FUNCTION_BLOCK Thomas_Object EXTENDS TcoCore.TcoObject
VAR
	_frank 		:	AKid_Object(THIS^);
	_andrew 	:	AKid_Object(THIS^);
	_christina 	:	AKid_Object(THIS^);
	_gianna 	:	AKid_Object(THIS^);
END_VAR

VAR
	_AskForTheFavor			:	AskForTheFavor_Task(THIS^);
END_VAR

METHOD AskForTheFavor : TcoCore.ITcoTask
VAR_INPUT
	Person_Requested 	:	REFERENCE TO Person_Object;
	RequestedFavor		:	STRING;
	ReturnFavor			:	STRING;
END_VAR
_AskForTheFavor(_Person_Requested := Person_Requested,_RequestedFavor :=RequestedFavor,_ReturnFavor:=ReturnFavor);

AskForTheFavor := _AskForTheFavor;
END_METHOD

END_FUNCTION_BLOCK

(* stored: Version 1.1.0.1, ProductVersion 3.1.4024.9
   POU Thomas_Object: Id {69d01a44-cebd-0fff-162d-7a59f62e3932}, SpecialFunc None
   Method AskForTheFavor: Id {c23a00a7-2858-0893-1a83-a9e7f9ad39a2} *)
